(* CODESYS project P_Active.xml

Project tree, tasks and I/O mapping:
*)

// P_Active
{attribute 'monitoring' := 'call'}
PROPERTY P_Active : BOOL
END_PROPERTY
